// LS Electric XG5000 project: test
// PLC LSPLC
// module base 0 slot 0: 입출력 모듈:XBC-DR32H (DC 24V 입력, 릴레이 출력 32점)

PROGRAM NewProgram (task: 스캔 프로그램)

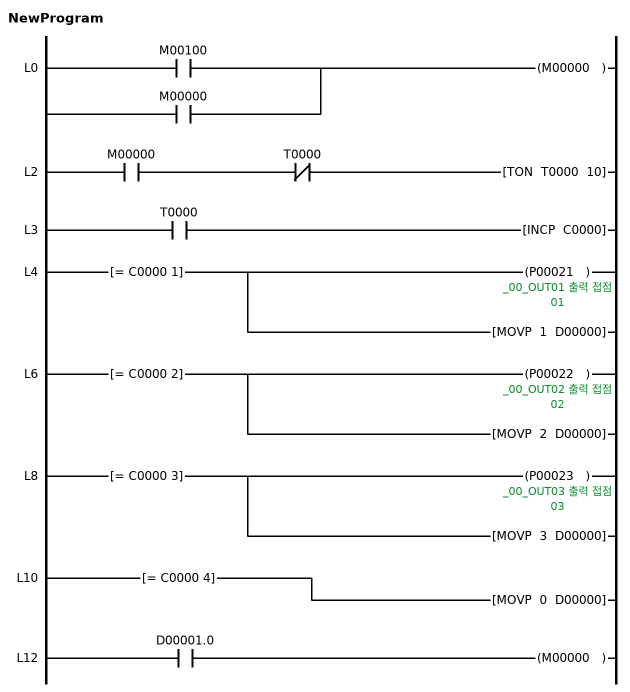
; L0
LOAD      M00100
OR        M00000
OUT       M00000
; L2
LOAD      M00000
AND NOT   T0000
TON       T0000 10
; L3
LOAD      T0000
INCP      C0000
; L4
LOAD=     C0000 1
OUT       P00021	// _00_OUT01 출력 접점 01
MOVP      1 D00000
; L6
LOAD=     C0000 2
OUT       P00022	// _00_OUT02 출력 접점 02
MOVP      2 D00000
; L8
LOAD=     C0000 3
OUT       P00023	// _00_OUT03 출력 접점 03
MOVP      3 D00000
; L10
LOAD=     C0000 4
MOVP      0 D00000
; L12
LOAD      D00001.0
OUT       M00000